Fanuc KAREL source: ko00035.KL

-- PROVISIONAL review KL for V1013-1; original PC SHA256 c9ddc7090b62394fb268791d6b4a43a1b53a0ff5f33ec1a8cfb098d569f88535
-- Incomplete behavior may be omitted. Consult companion uncertainty JSON. Do not deploy.
PROGRAM KO00035
%NOLOCKGROUP
BEGIN
  -- UNRESOLVED_PC offsets 5-12; opcodes 9D,23
  -- UNRESOLVED_PC offsets 17-66; opcodes 27,27,49,7E,AD,22,1C,22,31,7E,4A
  -- UNRESOLVED_PC offsets 71-75; opcodes 7F
END KO00035
